(* IEC 61131-3 sources: llm-plc-st-eval/data/definitivo/qwen2.5-coder_14b/C3/zero_shot, 3 files *)

(* ---- ejec_1.st ---- *)
```pascal
PROGRAM PRG_Conversion
VAR
    btnMarcha, btnParo : BOOL;  // Entradas
    motor, lampara : BOOL;      // Salidas
    T1 : TON;                   // Temporizador
END_VAR

// Rama 1: btnMarcha OR motor AND btnParo -> motor
motor := (btnMarcha OR motor) AND btnParo;

// Rama 2: motor -> T1 (10 segundos)
IF motor THEN
    T1(IN := TRUE, PT := T#10S);
ELSE
    T1(IN := FALSE);
END_IF;

// Rama 3: T1.Q -> lampara
lampara := T1.Q;
```

Este código en Structured Text (ST) implementa el comportamiento descrito en el Ladder Diagram, utilizando las variables y temporizadores especificados.

(* ---- ejec_2.st ---- *)
```pascal
PROGRAM PRG_Conversion
VAR
    btnMarcha, btnParo : BOOL;  // Entradas
    motor, lampara : BOOL;      // Salidas
    T1 : TON;                   // Temporizador
END_VAR

// Rama 1: btnMarcha OR motor AND btnParo -> motor
motor := (btnMarcha OR motor) AND btnParo;

// Rama 2: motor -> T1 (10 segundos)
IF motor THEN
    T1(IN := TRUE, PT := T#10S);
ELSE
    T1(IN := FALSE);
END_IF;

// Rama 3: T1.Q -> lampara
lampara := T1.Q;
```

Este código en Structured Text (ST) implementa el comportamiento descrito en el Ladder Diagram, utilizando las variables y temporizadores especificados.

(* ---- ejec_3.st ---- *)
```pascal
PROGRAM PRG_Conversion
VAR
    btnMarcha, btnParo : BOOL;  // Entradas
    motor, lampara : BOOL;      // Salidas
    T1 : TON;                   // Temporizador de 10 segundos
END_VAR

// Rama 1: btnMarcha y motor en paralelo, en serie con btnParo, alimentan motor
motor := (btnMarcha OR motor) AND btnParo;

// Rama 2: motor alimenta el temporizador T1 con tiempo preestablecido de 10 segundos
IF motor THEN
    T1(IN := TRUE, PT := T#10S);
ELSE
    T1(IN := FALSE);
END_IF;

// Rama 3: T1.Q alimenta la bobina lampara
lampara := T1.Q;
```

Este código en Structured Text (ST) cumple con el comportamiento descrito en el Ladder Diagram, utilizando las variables y temporizadores especificados.
